LAYER Default
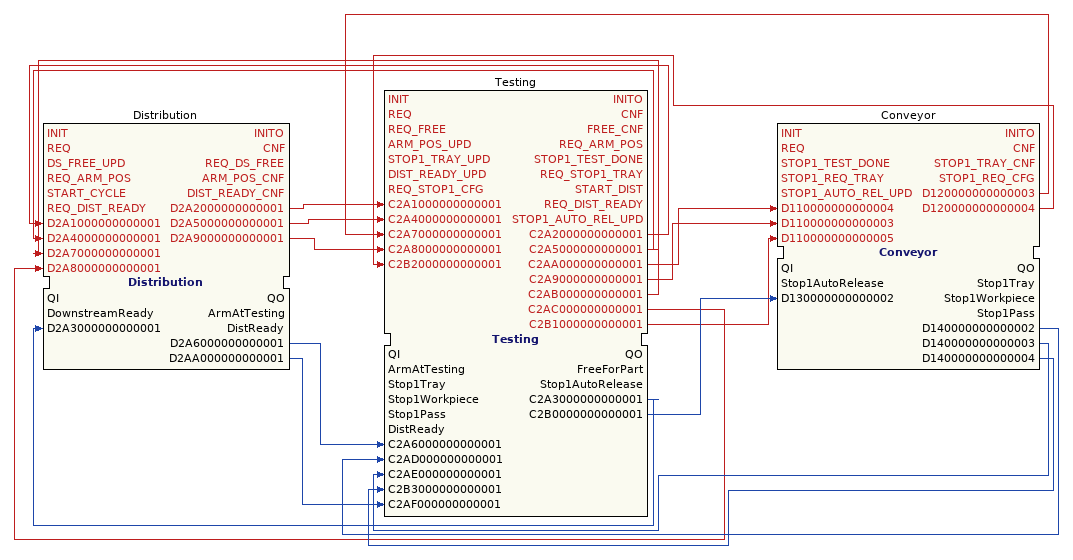
  FBS
    Distribution : Distribution;
    Testing : Testing;
    Conveyor : Conveyor;
  END_FBS
  EVENT_CONNECTIONS
    Testing.C2A2000000000001 TO Distribution.D2A1000000000001;
    Distribution.D2A2000000000001 TO Testing.C2A1000000000001;
    Distribution.D2A5000000000001 TO Testing.C2A4000000000001;
    Testing.C2A5000000000001 TO Distribution.D2A4000000000001;
    Conveyor.D120000000000003 TO Testing.C2A7000000000001;
    Testing.C2AA000000000001 TO Conveyor.D110000000000004;
    Testing.C2A9000000000001 TO Conveyor.D110000000000003;
    Testing.C2AB000000000001 TO Distribution.D2A7000000000001;
    Testing.C2AC000000000001 TO Distribution.D2A8000000000001;
    Distribution.D2A9000000000001 TO Testing.C2A8000000000001;
    Testing.C2B1000000000001 TO Conveyor.D110000000000005;
    Conveyor.D120000000000004 TO Testing.C2B2000000000001;
  END_CONNECTIONS
  DATA_CONNECTIONS
    Testing.C2A3000000000001 TO Distribution.D2A3000000000001;
    Distribution.D2A6000000000001 TO Testing.C2A6000000000001;
    Conveyor.D140000000000002 TO Testing.C2AD000000000001;
    Conveyor.D140000000000003 TO Testing.C2AE000000000001;
    Conveyor.D140000000000004 TO Testing.C2B3000000000001;
    Testing.C2B0000000000001 TO Conveyor.D130000000000002;
    Distribution.D2AA000000000001 TO Testing.C2AF000000000001;
  END_CONNECTIONS
END_LAYER
